// SIMATIC S7-200 project (STEP 7-Micro/WIN), CPU 226 CN REL 02.01

SYMBOL_TABLE USUARIO1
SP1              I0.0     // Sensor del tubo inferior
SP               I0.1     // Sensor del tubo superiro
SST              I0.2     // Sensor salida del tubo
SG               I0.3     // Sensor de recogida de pieza
SF               I0.4     // Sensor de posicion de pieza grande
SM1B             I0.5     // Sensor magnetico extendido del liberador
SM1A             I0.6     // Sensor magnetico retraido del liberador
SM2B             I0.7     // Sensor magnetico extendido del sujetador
SM2A             I1.0     // Sensor magnetico retraido del sujetador
SM3A             I1.1     // Sensor de giro antihorario
SM3B             I1.2     // Sensor de giro horario
SM6              I1.3     // Sensor de garra abierto
SM4B             I1.4     // Sensor magnetico extendido vertical
SM4A             I1.5     // Sensor magnetico retraido vertical
SM5A             I1.6     // Sensor magnetico retraido horizontal
SM5B             I1.7     // Sensor magnetico extendido horizontal
SB_2             I2.4     // Pulsador paro
SB_1             I2.5     // Pulsaodr de marcha
QS               I2.6     // Zeta de emergencia
SA               I2.7     // Selector de modo
KV2              Q0.0     // Cildro sujetador
KV1              Q0.1     // Cilindro liberador
KV3              Q0.2     // Cilindro rotatorio
KV6              Q0.3     // Cilindro de garra
KV4              Q0.4     // Cilindro vertical
KV5              Q0.5     // Cilindro horizontal
HL1B             Q0.7     // Baliza amarillo
HL2B             Q1.0     // Baliza verde
HL1              Q1.5     // Piloto amarillo
HL2              Q1.6     // Piloto verde
HL3              Q1.7     // Piloto rojo
E0               M0.0
E1               M0.1
E2               M0.2
E3               M0.3
E4               M0.4
E5               M0.5
E6               M0.6
E7               M0.7
E8               M1.0
E9               M1.1
E10              M1.2
E11              M1.3
E12              M1.4
E13              M1.5
E14              M1.6
EP               M1.7     // Paro momentaneo
EM               M2.0     // Estado  de emergencia
EM1              M2.1
END_SYMBOL_TABLE

ORGANIZATION_BLOCK PRINCIPAL:OB1
TITLE=COMENTARIOS DEL PROGRAMA
BEGIN
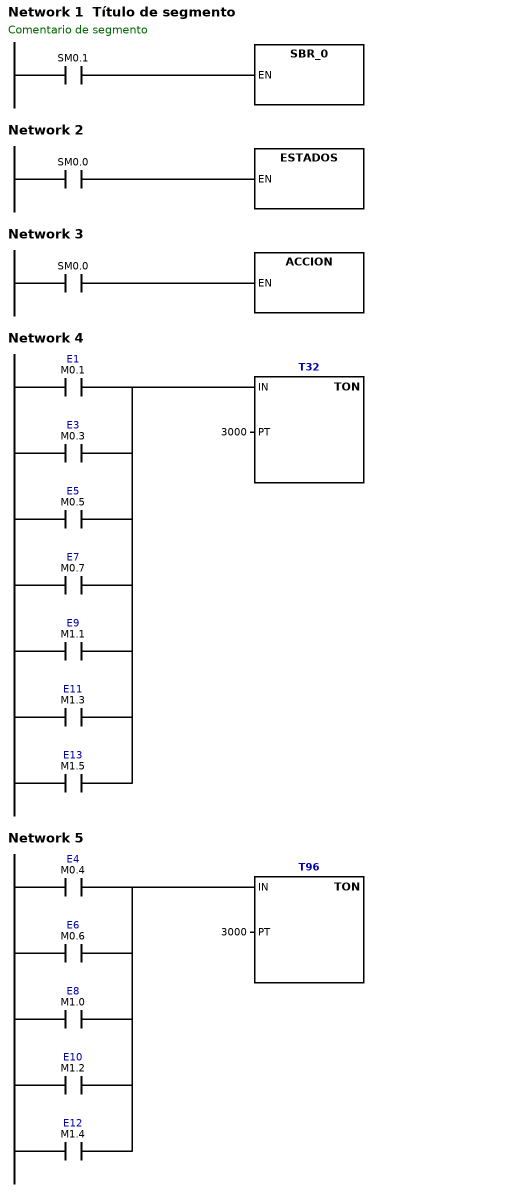
Network 1 // Título de segmento
// Comentario de segmento
LD     SM0.1
CALL   SBR_0:SBR0
Network 2
LD     SM0.0
CALL   ESTADOS:SBR1
Network 3
LD     SM0.0
CALL   ACCION:SBR2
Network 4
LD     E1:M0.1
O      E3:M0.3
O      E5:M0.5
O      E7:M0.7
O      E9:M1.1
O      E11:M1.3
O      E13:M1.5
TON    T32, 3000
Network 5
LD     E4:M0.4
O      E6:M0.6
O      E8:M1.0
O      E10:M1.2
O      E12:M1.4
TON    T96, 3000
END_ORGANIZATION_BLOCK

SUBROUTINE_BLOCK SBR_0:SBR0
TITLE=COMENTARIOS DE LA SUBRUTINA
BEGIN
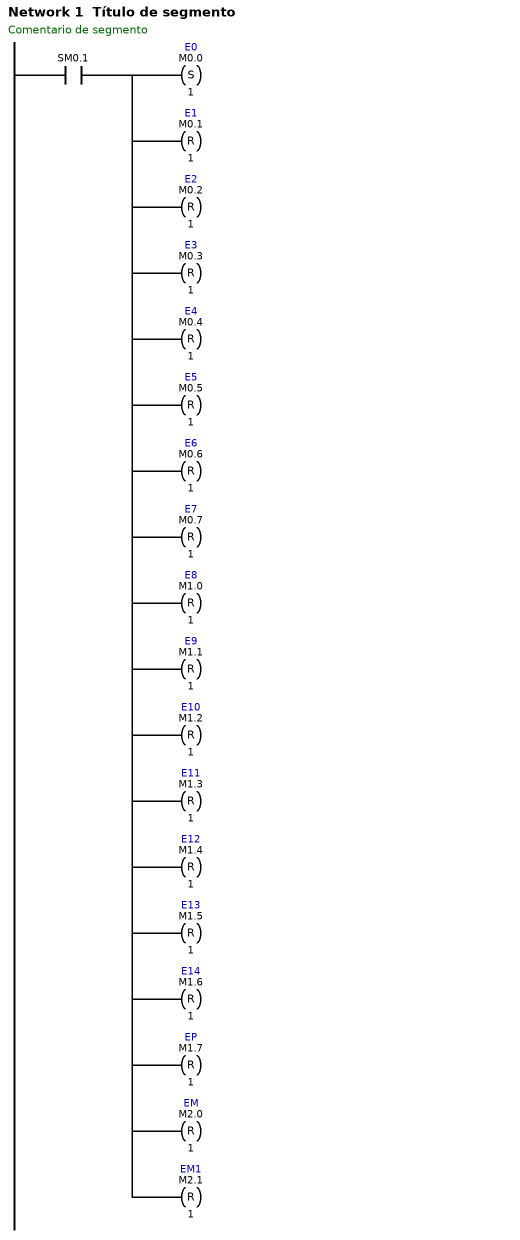
Network 1 // Título de segmento
// Comentario de segmento
LD     SM0.1
S      E0:M0.0, 1
R      E1:M0.1, 1
R      E2:M0.2, 1
R      E3:M0.3, 1
R      E4:M0.4, 1
R      E5:M0.5, 1
R      E6:M0.6, 1
R      E7:M0.7, 1
R      E8:M1.0, 1
R      E9:M1.1, 1
R      E10:M1.2, 1
R      E11:M1.3, 1
R      E12:M1.4, 1
R      E13:M1.5, 1
R      E14:M1.6, 1
R      EP:M1.7, 1
R      EM:M2.0, 1
R      EM1:M2.1, 1
END_SUBROUTINE_BLOCK

SUBROUTINE_BLOCK ESTADOS:SBR1
TITLE=COMENTARIOS DE LA SUBRUTINA
BEGIN
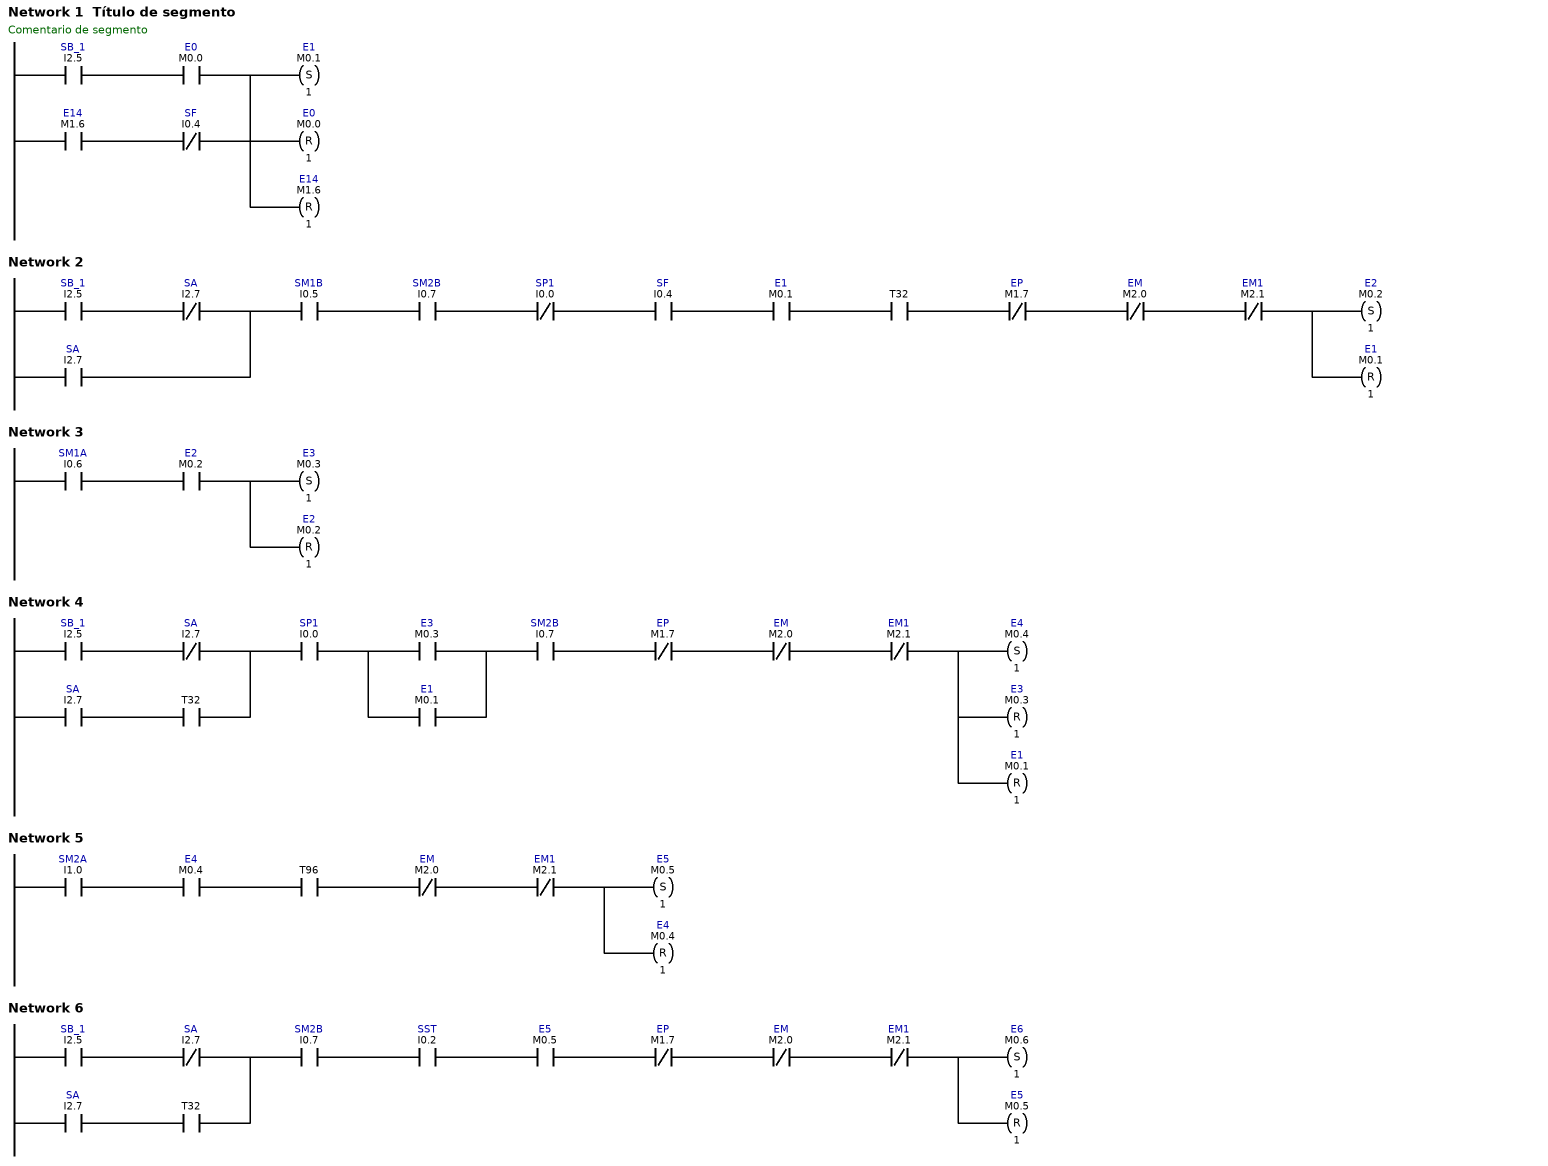
Network 1 // Título de segmento
// Comentario de segmento
LD     SB_1:I2.5
A      E0:M0.0
LD     E14:M1.6
AN     SF:I0.4
OLD
S      E1:M0.1, 1
R      E0:M0.0, 1
R      E14:M1.6, 1
Network 2
LD     SB_1:I2.5
AN     SA:I2.7
O      SA:I2.7
A      SM1B:I0.5
A      SM2B:I0.7
AN     SP1:I0.0
A      SF:I0.4
A      E1:M0.1
A      T32
AN     EP:M1.7
AN     EM:M2.0
AN     EM1:M2.1
S      E2:M0.2, 1
R      E1:M0.1, 1
Network 3
LD     SM1A:I0.6
A      E2:M0.2
S      E3:M0.3, 1
R      E2:M0.2, 1
Network 4
LD     SB_1:I2.5
AN     SA:I2.7
LD     SA:I2.7
A      T32
OLD
A      SP1:I0.0
LD     E3:M0.3
O      E1:M0.1
ALD
A      SM2B:I0.7
AN     EP:M1.7
AN     EM:M2.0
AN     EM1:M2.1
S      E4:M0.4, 1
R      E3:M0.3, 1
R      E1:M0.1, 1
Network 5
LD     SM2A:I1.0
A      E4:M0.4
A      T96
AN     EM:M2.0
AN     EM1:M2.1
S      E5:M0.5, 1
R      E4:M0.4, 1
Network 6
LD     SB_1:I2.5
AN     SA:I2.7
LD     SA:I2.7
A      T32
OLD
A      SM2B:I0.7
A      SST:I0.2
A      E5:M0.5
AN     EP:M1.7
AN     EM:M2.0
AN     EM1:M2.1
S      E6:M0.6, 1
R      E5:M0.5, 1
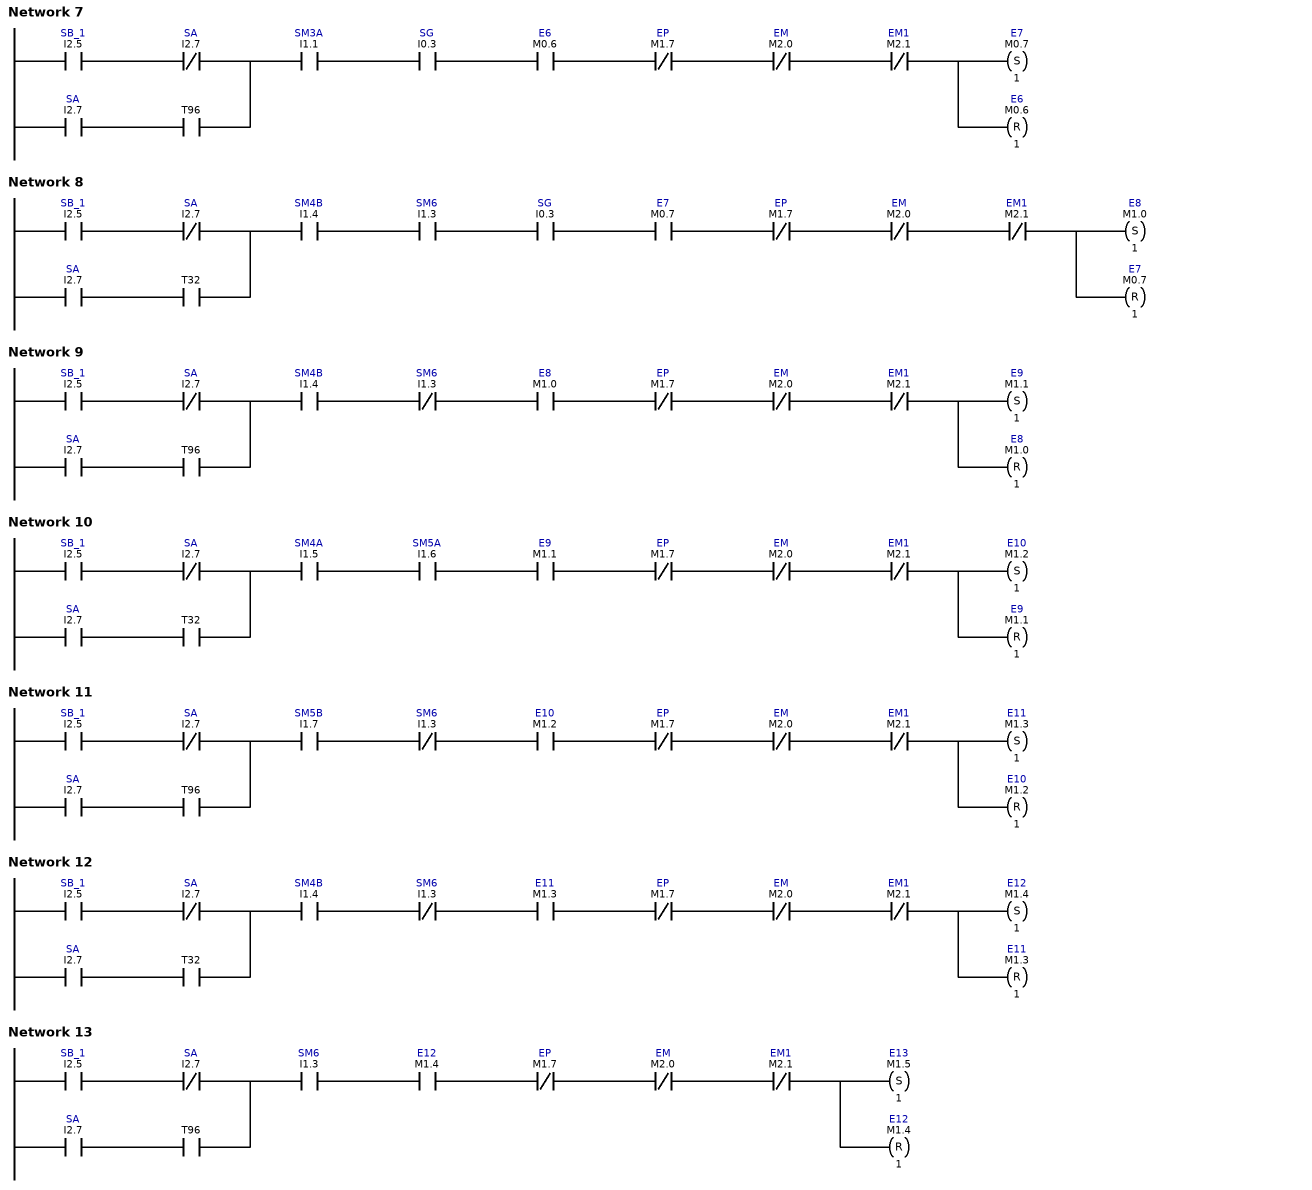
Network 7
LD     SB_1:I2.5
AN     SA:I2.7
LD     SA:I2.7
A      T96
OLD
A      SM3A:I1.1
A      SG:I0.3
A      E6:M0.6
AN     EP:M1.7
AN     EM:M2.0
AN     EM1:M2.1
S      E7:M0.7, 1
R      E6:M0.6, 1
Network 8
LD     SB_1:I2.5
AN     SA:I2.7
LD     SA:I2.7
A      T32
OLD
A      SM4B:I1.4
A      SM6:I1.3
A      SG:I0.3
A      E7:M0.7
AN     EP:M1.7
AN     EM:M2.0
AN     EM1:M2.1
S      E8:M1.0, 1
R      E7:M0.7, 1
Network 9
LD     SB_1:I2.5
AN     SA:I2.7
LD     SA:I2.7
A      T96
OLD
A      SM4B:I1.4
AN     SM6:I1.3
A      E8:M1.0
AN     EP:M1.7
AN     EM:M2.0
AN     EM1:M2.1
S      E9:M1.1, 1
R      E8:M1.0, 1
Network 10
LD     SB_1:I2.5
AN     SA:I2.7
LD     SA:I2.7
A      T32
OLD
A      SM4A:I1.5
A      SM5A:I1.6
A      E9:M1.1
AN     EP:M1.7
AN     EM:M2.0
AN     EM1:M2.1
S      E10:M1.2, 1
R      E9:M1.1, 1
Network 11
LD     SB_1:I2.5
AN     SA:I2.7
LD     SA:I2.7
A      T96
OLD
A      SM5B:I1.7
AN     SM6:I1.3
A      E10:M1.2
AN     EP:M1.7
AN     EM:M2.0
AN     EM1:M2.1
S      E11:M1.3, 1
R      E10:M1.2, 1
Network 12
LD     SB_1:I2.5
AN     SA:I2.7
LD     SA:I2.7
A      T32
OLD
A      SM4B:I1.4
AN     SM6:I1.3
A      E11:M1.3
AN     EP:M1.7
AN     EM:M2.0
AN     EM1:M2.1
S      E12:M1.4, 1
R      E11:M1.3, 1
Network 13
LD     SB_1:I2.5
AN     SA:I2.7
LD     SA:I2.7
A      T96
OLD
A      SM6:I1.3
A      E12:M1.4
AN     EP:M1.7
AN     EM:M2.0
AN     EM1:M2.1
S      E13:M1.5, 1
R      E12:M1.4, 1
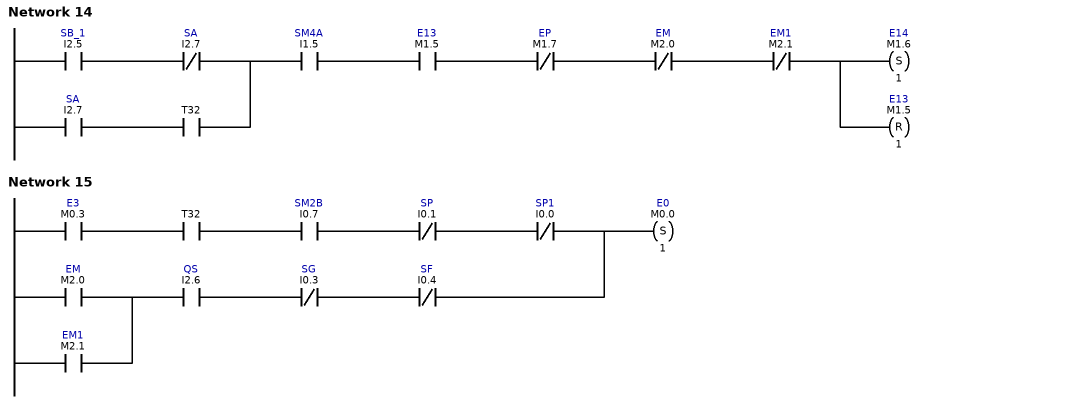
Network 14
LD     SB_1:I2.5
AN     SA:I2.7
LD     SA:I2.7
A      T32
OLD
A      SM4A:I1.5
A      E13:M1.5
AN     EP:M1.7
AN     EM:M2.0
AN     EM1:M2.1
S      E14:M1.6, 1
R      E13:M1.5, 1
Network 15
LD     E3:M0.3
A      T32
A      SM2B:I0.7
AN     SP:I0.1
AN     SP1:I0.0
LD     EM:M2.0
O      EM1:M2.1
A      QS:I2.6
AN     SG:I0.3
AN     SF:I0.4
OLD
S      E0:M0.0, 1
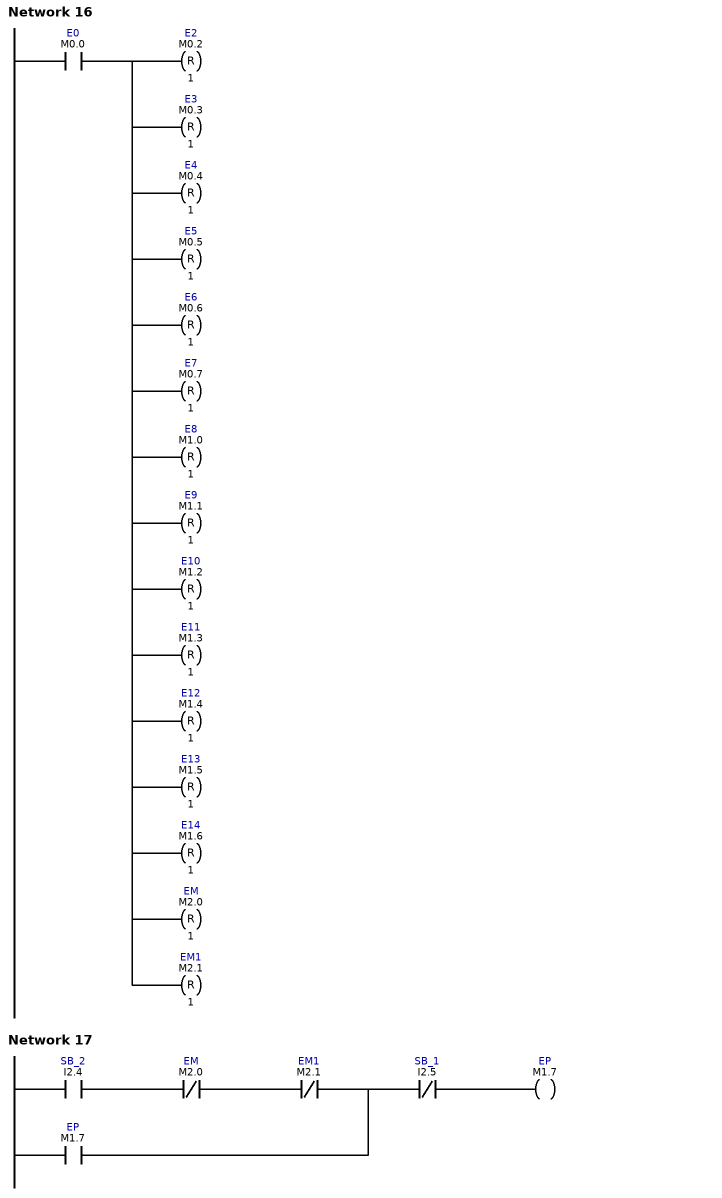
Network 16
LD     E0:M0.0
R      E2:M0.2, 1
R      E3:M0.3, 1
R      E4:M0.4, 1
R      E5:M0.5, 1
R      E6:M0.6, 1
R      E7:M0.7, 1
R      E8:M1.0, 1
R      E9:M1.1, 1
R      E10:M1.2, 1
R      E11:M1.3, 1
R      E12:M1.4, 1
R      E13:M1.5, 1
R      E14:M1.6, 1
R      EM:M2.0, 1
R      EM1:M2.1, 1
Network 17
LD     SB_2:I2.4
AN     EM:M2.0
AN     EM1:M2.1
O      EP:M1.7
AN     SB_1:I2.5
=      EP:M1.7
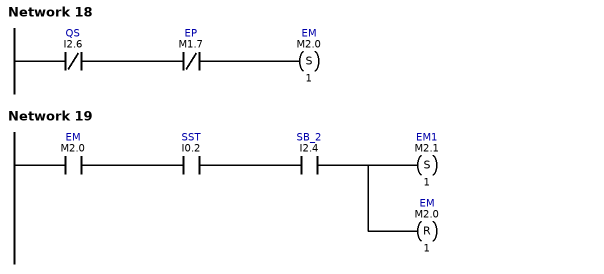
Network 18
LDN    QS:I2.6
AN     EP:M1.7
S      EM:M2.0, 1
Network 19
LD     EM:M2.0
A      SST:I0.2
A      SB_2:I2.4
S      EM1:M2.1, 1
R      EM:M2.0, 1
END_SUBROUTINE_BLOCK

SUBROUTINE_BLOCK ACCION:SBR2
TITLE=COMENTARIOS DE LA SUBRUTINA
BEGIN
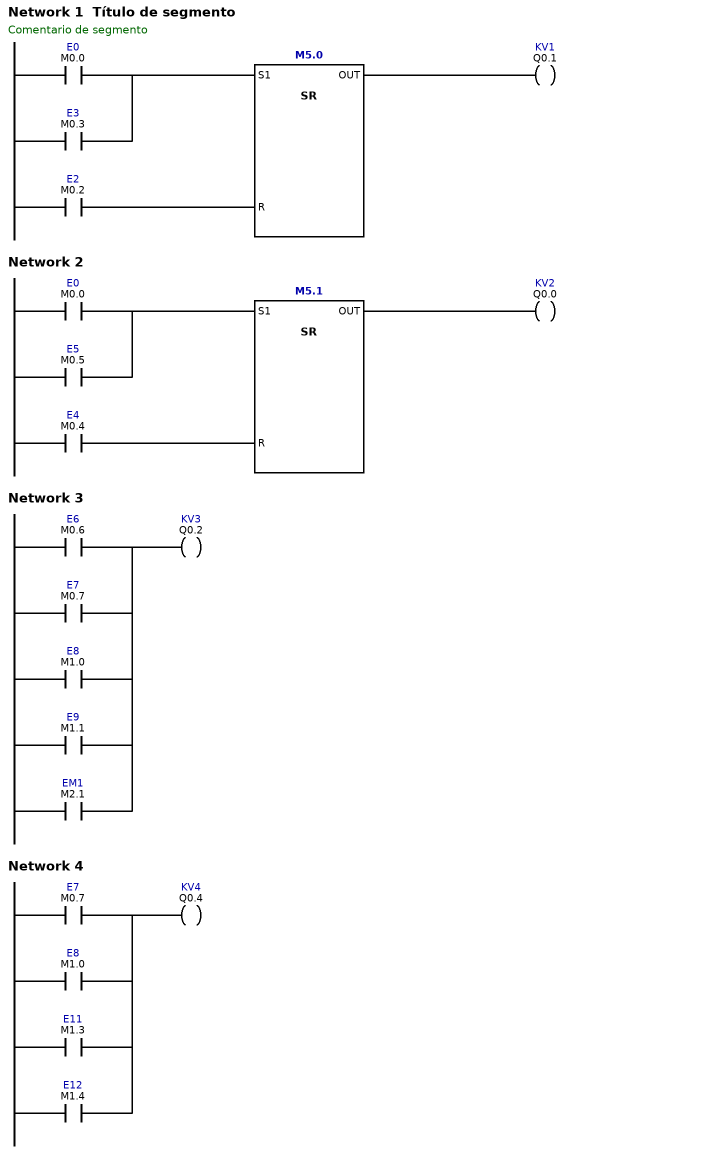
Network 1 // Título de segmento
// Comentario de segmento
LD     E0:M0.0
O      E3:M0.3
LD     E2:M0.2
NOT
A      M5.0
OLD
=      M5.0
=      KV1:Q0.1
Network 2
LD     E0:M0.0
O      E5:M0.5
LD     E4:M0.4
NOT
A      M5.1
OLD
=      M5.1
=      KV2:Q0.0
Network 3
LD     E6:M0.6
O      E7:M0.7
O      E8:M1.0
O      E9:M1.1
O      EM1:M2.1
=      KV3:Q0.2
Network 4
LD     E7:M0.7
O      E8:M1.0
O      E11:M1.3
O      E12:M1.4
=      KV4:Q0.4
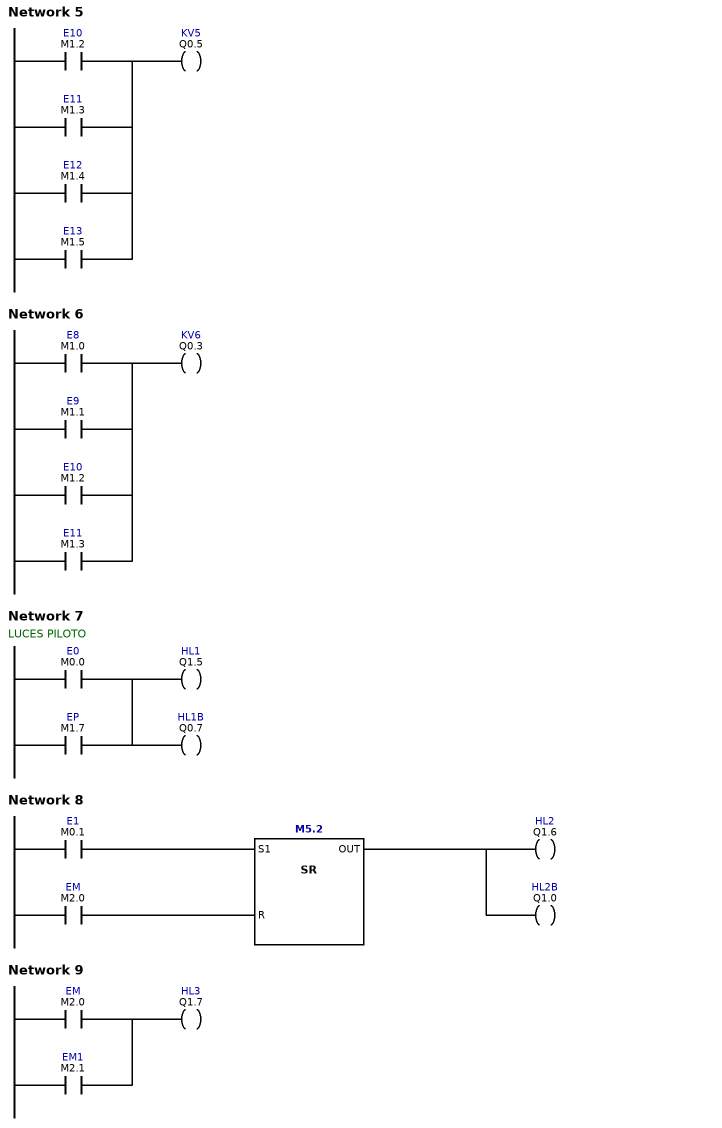
Network 5
LD     E10:M1.2
O      E11:M1.3
O      E12:M1.4
O      E13:M1.5
=      KV5:Q0.5
Network 6
LD     E8:M1.0
O      E9:M1.1
O      E10:M1.2
O      E11:M1.3
=      KV6:Q0.3
Network 7
// LUCES PILOTO
LD     E0:M0.0
O      EP:M1.7
=      HL1:Q1.5
=      HL1B:Q0.7
Network 8
LD     E1:M0.1
LD     EM:M2.0
NOT
A      M5.2
OLD
=      M5.2
=      HL2:Q1.6
=      HL2B:Q1.0
Network 9
LD     EM:M2.0
O      EM1:M2.1
=      HL3:Q1.7
END_SUBROUTINE_BLOCK
